RoboDK station: XARM5.rdk

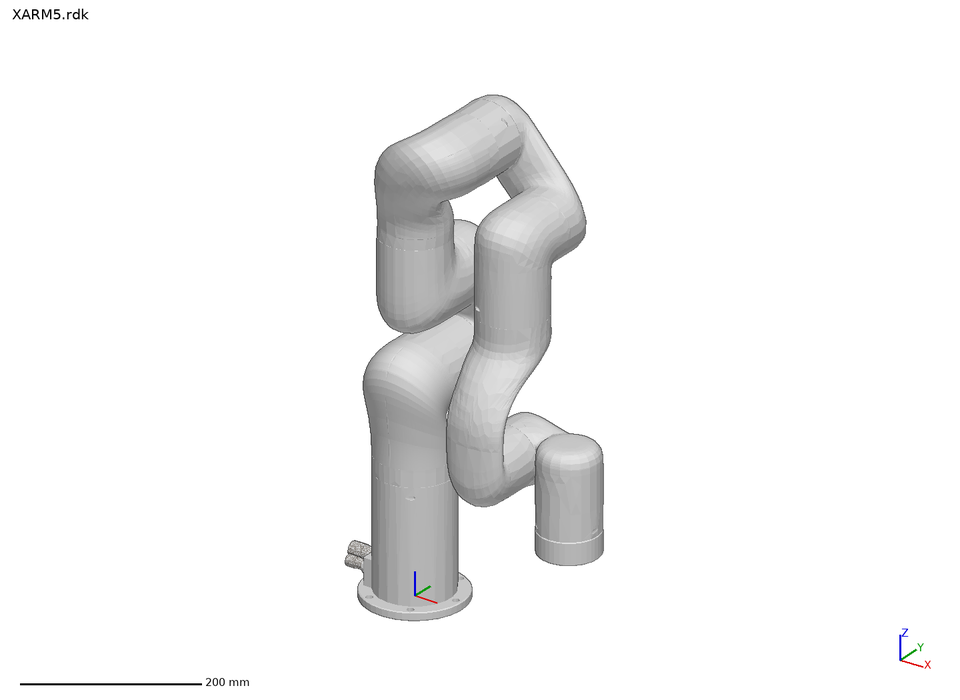
[picture v0: the station drawn from its stored meshes, robots at their saved joint values, targets as dots, program paths as lines]
Station XARM5 (saved by RoboDK 6.2.0). Poses are relative to the parent item; angles as X-Y-Z fixed-axis rotations.
  - frame uFactory xArm5 Base at (0, 0, 0) mm
    - robot uFactory xArm5: 6 axes, payload 3 kg, reach 700 mm, repeatability 0.1 mm, weight 11.2 kg
        modified DH rows (alpha deg, a mm, theta deg, d mm): 0, 0, 0, 267; -90, 0, -79.35, 0; 0, 289.489, 79.35, 0; -90, 77.5, 0, 342.5; 90, 0, 0, 0; -90, 76, 0, 97
        joint limits [-360, -118, -225, -0.01, -97, -360] to [360, 120, 11, 0.01, 180, 360]; home [0, 0, 0, 0, 0, 0]; saved at [0, 0, 0, 0, 0, 0]
